Fanuc KAREL source: KD00055.KL

PROGRAM KD00055
%NOLOCKGROUP
VAR
  I: INTEGER
  J: INTEGER
  B: BOOLEAN
  R: REAL
  S: STRING[80]
BEGIN
  CONDITION[1]:
  WHEN DIN[1] = ON DO
    DOUT[2] = ON
  ENDCONDITION
END KD00055
